// TIA Portal V21 export
// export: Created 2026-08-21T20:18:54.2707311Z, ExportSetting None, DisplayName Totally Integrated Automation Portal, DisplayVersion V21, DisplayName STEP 7 Professional, DisplayVersion V21, DisplayName STEP 7 Safety, DisplayVersion V21, DisplayName Tech WebApplication, DisplayVersion V21, DisplayName WinCC Basic/Comfort/Advanced, DisplayVersion V21, DisplayName WinCC Professional, DisplayVersion V21, DisplayName WinCC Unified, DisplayVersion V21
TYPE "UDT_MTP_Procedure"
   STRUCT
      IsSelfCompleting : Bool;   // 1:Procedure Self-Completing; 0:Procedure Not Self-Completing
      ProcedureID : DWord;   // Procedure ID
      IsDefault : Bool;   // 1:Default procedure; 0:Not Default Procedure
   END_STRUCT;
END_TYPE
